Universal Robots PolyScope program: pick_and_place.urp

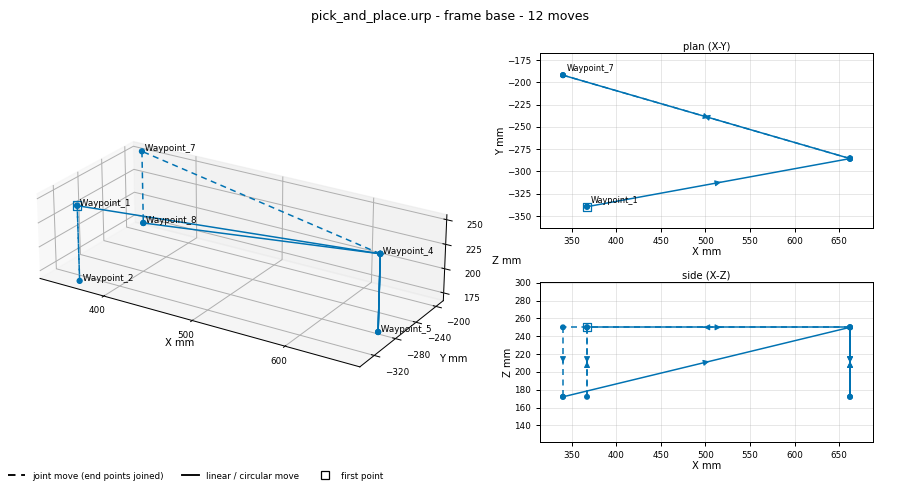
[picture p0: tool path of pick_and_place.urp in frame base, 12 of 12 moves have a stored position in this frame; points joined in program order, loops and branches not executed]
Program pick_and_place (installation=default directory=/ursim/programs/actividad 3 createdIn=3.15.8.106339 lastSavedIn=3.15.8.106339 robotSerialNumber=2018359999)
Calibrated DH parameters: a=[0, -0.425, -0.39225, 0, 0, 0]; d=[0.089159, 0, 0, 0.10915, 0.09465, 0.0823]; alpha=[1.570796, 0, 0, 1.570796, -1.570796, 0]; deltaTheta=[0, 0, 0, 0, 0, 0]
Robot Program (runOnlyOnce=false)
  Popup Message (haltProgram=false message=ENCENDER ENTRADA DIGITAL 0 inputType=Text)
  Wait DigitalInput pin=digital_in[0]; digitalValue=0
  MoveJ speed 60 deg/s, acceleration 80 deg/s^2 (useActiveTCP=true)
    Waypoint Waypoint_1: TCP in base x=367.081 y=-339.488 z=250 mm, rx=-0.0012 ry=3.1163 rz=0.0389 rad; joints [-30.485, -96.06, -111.318, -62.11, 91.961, 59.479] deg
    Waypoint Waypoint_2: TCP in base x=367.081 y=-339.488 z=172 mm, rx=-0.0012 ry=3.1163 rz=0.0389 rad; joints [-30.485, -102.442, -117.3, -49.747, 91.961, 59.479] deg
    Set DigitalOutput pin=digital_out[0]; digitalValue=0
    Wait Sleep waitTime=1
    Waypoint Waypoint_3: TCP in base x=367.081 y=-339.488 z=250 mm, rx=-0.0012 ry=3.1163 rz=0.0389 rad; joints [-30.485, -96.06, -111.318, -62.11, 91.961, 59.479] deg
  MoveL speed 250 mm/s, acceleration 1200 mm/s^2 (useActiveTCP=true) feature=Base
    Waypoint Waypoint_4: TCP in base x=662.184 y=-285.504 z=250 mm, rx=-0.0012 ry=3.1163 rz=0.0389 rad; joints [-14.82, -124.434, -71.721, -72.823, 91.75, 75.151] deg
    Waypoint Waypoint_5: TCP in base x=662.184 y=-285.504 z=172 mm, rx=-0.0012 ry=3.1163 rz=0.0389 rad; joints [-14.82, -128.33, -77.353, -63.295, 91.75, 75.151] deg
    Set DigitalOutput pin=digital_out[0]; digitalValue=1
    Wait Sleep waitTime=1
    Waypoint Waypoint_6: TCP in base x=662.184 y=-285.504 z=250 mm, rx=-0.0012 ry=3.1163 rz=0.0389 rad; joints [-14.82, -124.434, -71.721, -72.823, 91.75, 75.151] deg
  MoveJ speed 60 deg/s, acceleration 80 deg/s^2 (useActiveTCP=true)
    Waypoint Waypoint_7: TCP in base x=340.089 y=-191.936 z=250 mm, rx=-0.0012 ry=3.1163 rz=0.0389 rad; joints [-13.587, -80.504, -126.456, -61.979, 91.728, 76.384] deg
    Waypoint Waypoint_8: TCP in base x=340.089 y=-191.936 z=172 mm, rx=-0.0012 ry=3.1163 rz=0.0389 rad; joints [-13.587, -88.262, -133.542, -47.136, 91.728, 76.384] deg
    Set DigitalOutput pin=digital_out[0]; digitalValue=0
    Wait Sleep waitTime=1
    Waypoint Waypoint_9: TCP in base x=340.089 y=-191.936 z=172 mm, rx=-0.0012 ry=3.1163 rz=0.0389 rad; joints [-13.587, -88.262, -133.542, -47.136, 91.728, 76.384] deg
  MoveL speed 250 mm/s, acceleration 1200 mm/s^2 (useActiveTCP=true) feature=Base
    Waypoint Waypoint_10: TCP in base x=662.184 y=-285.504 z=250 mm, rx=-0.0012 ry=3.1163 rz=0.0389 rad; joints [-14.82, -124.434, -71.721, -72.823, 91.75, 75.151] deg
    Waypoint Waypoint_11: TCP in base x=662.184 y=-285.504 z=172 mm, rx=-0.0012 ry=3.1163 rz=0.0389 rad; joints [-14.82, -128.33, -77.353, -63.295, 91.75, 75.151] deg
    Set DigitalOutput pin=digital_out[0]; digitalValue=1
    Wait Sleep waitTime=1
    Waypoint Waypoint_12: TCP in base x=662.184 y=-285.504 z=250 mm, rx=-0.0012 ry=3.1163 rz=0.0389 rad; joints [-14.82, -124.434, -71.721, -72.823, 91.75, 75.151] deg
